(* IEC 61131-3 sources: plcassist-cli/packages/volt-lsp-iec/test-corpus/awa-palletizer/Device/Plc Logic/Application/Library Manager/(unresolved)/syssem interfaces, 1 file *)

(* ---- GVL.gvl ---- *)
VAR_GLOBAL
	SYSSEM_INVALID_HANDLE : UDINT := 16#FFFFFFFF;
END_VAR
